(* PLC project Geraetebeschreibungen, CODESYS CODESYS V3.5 SP21, author synthetisch *)
(* stored: creationDateTime 2026-10-31T10:00:00.0000000, version 1.0.0.0, modificationDateTime 2026-10-31T09:59:00.0000000, organization Comquent GmbH *)

CONFIGURATION Steuerung
  RESOURCE Application ON PLC
  END_RESOURCE
END_CONFIGURATION

CONFIGURATION I2C_Mux
END_CONFIGURATION

CONFIGURATION Expander
END_CONFIGURATION

CONFIGURATION Lichtsensor
END_CONFIGURATION
